Yaskawa INFORM job: PAT_CR.JBI

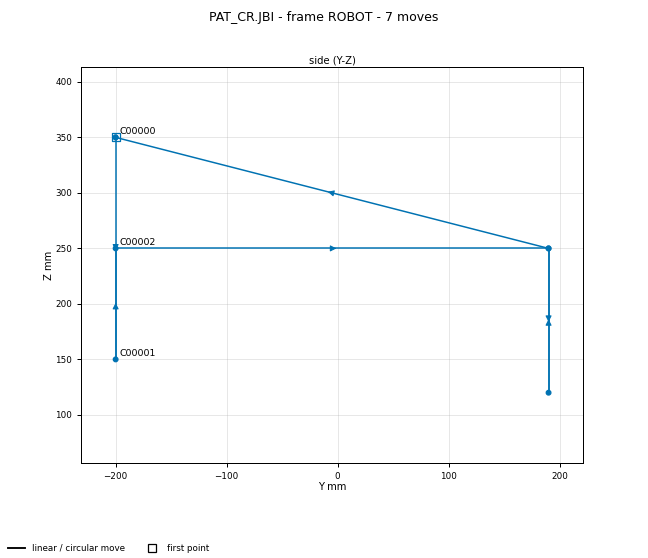
[picture p0: tool path of PAT_CR.JBI in frame ROBOT, 7 of 7 moves have a stored position in this frame; points joined in program order, loops and branches not executed]
/JOB
//NAME PAT_CR
//POS
///NPOS 7,0,0,0,0,0
///TOOL 0
///POSTYPE ROBOT
///RECTAN
///RCONF 0,0,0,0,0,0,0,0
C00000=450.000,-200.000,350.000,180.00,0.00,0.00
C00001=450.000,-200.000,150.000,180.00,0.00,0.00
C00002=450.000,-200.000,250.000,180.00,0.00,0.00
C00003=450.000,190.000,250.000,180.00,0.00,0.00
C00004=450.000,190.000,120.000,180.00,0.00,0.00
C00005=450.000,190.000,250.000,180.00,0.00,0.00
C00006=450.000,-200.000,350.000,180.00,0.00,0.00
//INST
///DATE 2026/11/02 14:40
///ATTR SC,RW
///GROUP1 RB1
NOP
'SYNTHETIC TEST DATA - NOT A REAL ROBOT JOB
MOVL C00000 V=200.0
MOVL C00001 V=80.0
DOUT OT#(1) ON
TIMER T=0.50
MOVL C00002 V=80.0 CR=10.0
MOVL C00003 V=250.0
MOVL C00004 V=80.0
TIMER T=3.00
DOUT OT#(1) OFF
TIMER T=0.50
MOVL C00005 V=80.0
MOVL C00006 V=200.0
END
